Staubli VAL3: _CalpCircle.pgx

program _CalpCircle(pointRs x_p1, pointRs x_p2, pointRs x_p3, pointRs& x_pCenter, bool& x_bStatus)
  local num x1
  local num y1
  local num x2
  local num y2
  local num x3
  local num y3
  local frame l_fFrame
  local num l_nFrameStatus
  local pointRs l_p3
  local pointRs l_p2
  local pointRs l_p1
  local pointRs l_pCenter
begin
  //圆心算法
  link(l_fFrame,world)
  l_nFrameStatus=setFrame(x_p1,x_p2,x_p3,l_fFrame)
  if l_nFrameStatus!=0
    //3点共线或任意2点过于接近
    popUpMsg("Error!!")
    x_bStatus=false
    return
  endIf
  link(l_p1,l_fFrame)
  link(l_p2,l_fFrame)
  link(l_p3,l_fFrame)
  l_p1.trsf=position(x_p1,l_fFrame)
  l_p2.trsf=position(x_p2,l_fFrame)
  l_p3.trsf=position(x_p3,l_fFrame)
  //
  x1=l_p1.trsf.x
  y1=l_p1.trsf.y
  x2=l_p2.trsf.x
  y2=l_p2.trsf.y
  x3=l_p3.trsf.x
  y3=l_p3.trsf.y
  //
  if((x3-x1)*(y2-y1)-(x2-x1)*(y3-y1))!=0
    link(l_pCenter,l_fFrame)
    l_pCenter.trsf={0,0,0,0,0,0}
    l_pCenter.trsf.x=((y2-y1)*(y3*y3-y1*y1+x3*x3-x1*x1)-(y3-y1)*(y2*y2-y1*y1+x2*x2-x1*x1))/(2*(x3-x1)*(y2-y1)-2*(x2-x1)*(y3-y1))
    l_pCenter.trsf.y=((x2-x1)*(x3*x3-x1*x1+y3*y3-y1*y1)-(x3-x1)*(x2*x2-x1*x1+y2*y2-y1*y1))/(2*(y3-y1)*(x2-x1)-2*(y2-y1)*(x3-x1))
    x_pCenter.trsf=position(l_pCenter,world)
    x_bStatus=true
  else
    x_bStatus=false
    return
 endIf
end
